SYSTEM PID_Basic_Adaptive (* Minimal synthetic PID with one direct gain update; native validation pending *)
  APPLICATION Basic_Control (* Process, identifier/tuner and flag PID *)
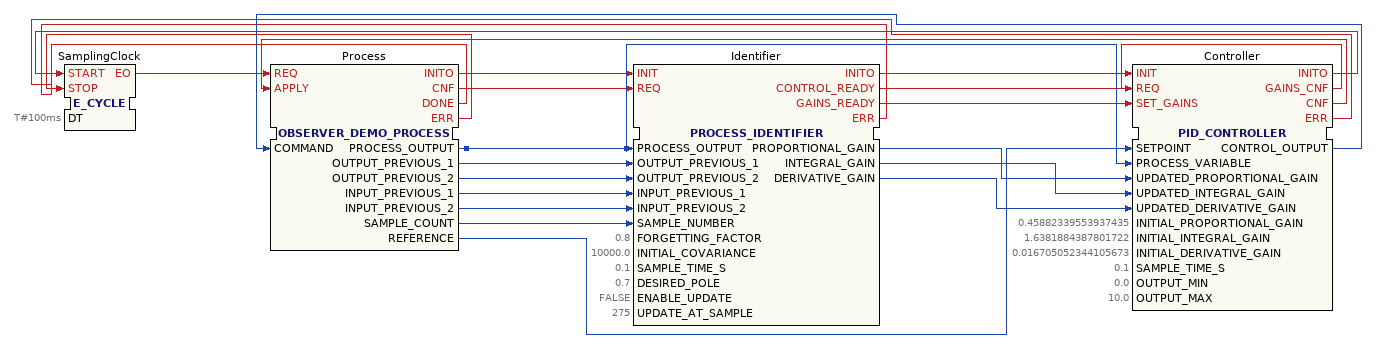
    FBS
      SamplingClock : E_CYCLE(DT := T#100ms);
      Process : OBSERVER_DEMO_PROCESS;
      Identifier : PROCESS_IDENTIFIER(FORGETTING_FACTOR := 0.8, INITIAL_COVARIANCE := 10000.0, SAMPLE_TIME_S := 0.1, DESIRED_POLE := 0.7, ENABLE_UPDATE := FALSE, UPDATE_AT_SAMPLE := 275);
      Controller : PID_CONTROLLER(INITIAL_PROPORTIONAL_GAIN := 0.45882339553937435, INITIAL_INTEGRAL_GAIN := 1.6381884387801722, INITIAL_DERIVATIVE_GAIN := 0.016705052344105673, SAMPLE_TIME_S := 0.1, OUTPUT_MIN := 0.0, OUTPUT_MAX := 10.0);
    END_FBS
    EVENT_CONNECTIONS
      Process.INITO TO Identifier.INIT;
      Identifier.INITO TO Controller.INIT;
      Controller.INITO TO SamplingClock.START;
      SamplingClock.EO TO Process.REQ;
      Process.CNF TO Identifier.REQ;
      Identifier.CONTROL_READY TO Controller.REQ;
      Identifier.GAINS_READY TO Controller.SET_GAINS;
      Controller.GAINS_CNF TO Controller.REQ;
      Controller.CNF TO Process.APPLY;
      Process.DONE TO SamplingClock.STOP;
      Process.ERR TO SamplingClock.STOP;
      Identifier.ERR TO SamplingClock.STOP;
      Controller.ERR TO SamplingClock.STOP;
    END_CONNECTIONS
    DATA_CONNECTIONS
      Process.PROCESS_OUTPUT TO Identifier.PROCESS_OUTPUT;
      Process.OUTPUT_PREVIOUS_1 TO Identifier.OUTPUT_PREVIOUS_1;
      Process.OUTPUT_PREVIOUS_2 TO Identifier.OUTPUT_PREVIOUS_2;
      Process.INPUT_PREVIOUS_1 TO Identifier.INPUT_PREVIOUS_1;
      Process.INPUT_PREVIOUS_2 TO Identifier.INPUT_PREVIOUS_2;
      Process.SAMPLE_COUNT TO Identifier.SAMPLE_NUMBER;
      Process.REFERENCE TO Controller.SETPOINT;
      Process.PROCESS_OUTPUT TO Controller.PROCESS_VARIABLE;
      Controller.CONTROL_OUTPUT TO Process.COMMAND;
      Identifier.PROPORTIONAL_GAIN TO Controller.UPDATED_PROPORTIONAL_GAIN;
      Identifier.INTEGRAL_GAIN TO Controller.UPDATED_INTEGRAL_GAIN;
      Identifier.DERIVATIVE_GAIN TO Controller.UPDATED_DERIVATIVE_GAIN;
    END_CONNECTIONS
  END_APPLICATION
  DEVICE LocalObserver : FORTE_PC(MGR_ID := "localhost:61499") (* Local synthetic test only *)
    {SET_ATTRIBUTE(Profile, HOLOBLOC)}
    RESOURCE EMB_RES : EMB_RES
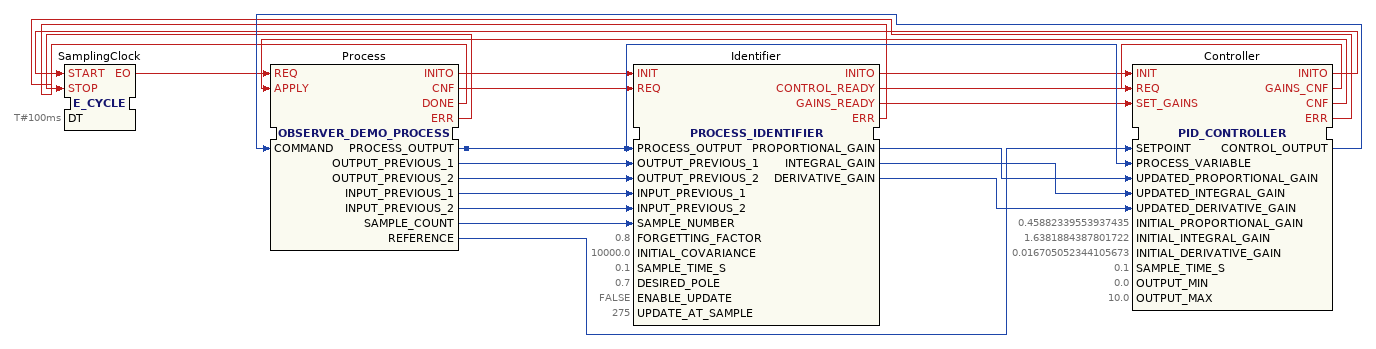
      FBS
        SamplingClock : E_CYCLE(DT := T#100ms);
        Process : OBSERVER_DEMO_PROCESS;
        Identifier : PROCESS_IDENTIFIER(FORGETTING_FACTOR := 0.8, INITIAL_COVARIANCE := 10000.0, SAMPLE_TIME_S := 0.1, DESIRED_POLE := 0.7, ENABLE_UPDATE := FALSE, UPDATE_AT_SAMPLE := 275);
        Controller : PID_CONTROLLER(INITIAL_PROPORTIONAL_GAIN := 0.45882339553937435, INITIAL_INTEGRAL_GAIN := 1.6381884387801722, INITIAL_DERIVATIVE_GAIN := 0.016705052344105673, SAMPLE_TIME_S := 0.1, OUTPUT_MIN := 0.0, OUTPUT_MAX := 10.0);
      END_FBS
      EVENT_CONNECTIONS
        Process.INITO TO Identifier.INIT;
        Identifier.INITO TO Controller.INIT;
        Controller.INITO TO SamplingClock.START;
        SamplingClock.EO TO Process.REQ;
        Process.CNF TO Identifier.REQ;
        Identifier.CONTROL_READY TO Controller.REQ;
        Identifier.GAINS_READY TO Controller.SET_GAINS;
        Controller.GAINS_CNF TO Controller.REQ;
        Controller.CNF TO Process.APPLY;
        Process.DONE TO SamplingClock.STOP;
        Process.ERR TO SamplingClock.STOP;
        Identifier.ERR TO SamplingClock.STOP;
        Controller.ERR TO SamplingClock.STOP;
      END_CONNECTIONS
      DATA_CONNECTIONS
        Process.PROCESS_OUTPUT TO Identifier.PROCESS_OUTPUT;
        Process.OUTPUT_PREVIOUS_1 TO Identifier.OUTPUT_PREVIOUS_1;
        Process.OUTPUT_PREVIOUS_2 TO Identifier.OUTPUT_PREVIOUS_2;
        Process.INPUT_PREVIOUS_1 TO Identifier.INPUT_PREVIOUS_1;
        Process.INPUT_PREVIOUS_2 TO Identifier.INPUT_PREVIOUS_2;
        Process.SAMPLE_COUNT TO Identifier.SAMPLE_NUMBER;
        Process.REFERENCE TO Controller.SETPOINT;
        Process.PROCESS_OUTPUT TO Controller.PROCESS_VARIABLE;
        Controller.CONTROL_OUTPUT TO Process.COMMAND;
        Identifier.PROPORTIONAL_GAIN TO Controller.UPDATED_PROPORTIONAL_GAIN;
        Identifier.INTEGRAL_GAIN TO Controller.UPDATED_INTEGRAL_GAIN;
        Identifier.DERIVATIVE_GAIN TO Controller.UPDATED_DERIVATIVE_GAIN;
      END_CONNECTIONS
    END_RESOURCE
  END_DEVICE
  MAPPINGS
    Basic_Control.SamplingClock ON LocalObserver.EMB_RES.SamplingClock;
    Basic_Control.Process ON LocalObserver.EMB_RES.Process;
    Basic_Control.Identifier ON LocalObserver.EMB_RES.Identifier;
    Basic_Control.Controller ON LocalObserver.EMB_RES.Controller;
  END_MAPPINGS
END_SYSTEM
